(* PLC project Vn_networks5, Beckhoff Automation GmbH TwinCAT PLC Control 3.5.13.21 *)
(* stored: creationDateTime 1970-01-01T00:00:00 *)

PROGRAM Vn_networks5

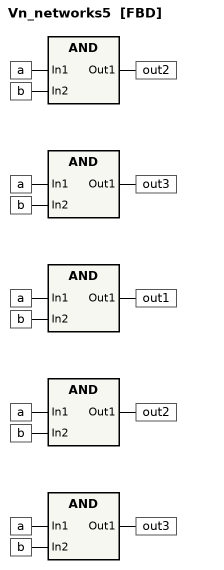
(* FBD diagram, written out as Structured Text *)
out2 := a AND b;
out3 := a AND b;
out1 := a AND b;
out2 := a AND b;
out3 := a AND b;
END_PROGRAM
